Fanuc KAREL source: KA00095.KL

PROGRAM KA00095
%NOLOCKGROUP
VAR
  SRC: JOINTPOS
  DST: ARRAY[2] OF BYTE
BEGIN
  DST[1] = SRC
END KA00095
